Fanuc KAREL source: KC00004.KL

PROGRAM KC00004
%NOLOCKGROUP
%ENVIRONMENT PC
VAR
  I: INTEGER
  J: INTEGER
  K: INTEGER
  R: REAL
  B: BOOLEAN
  S: STRING[80]
  T: STRING[80]
  P: PATH
  Q: PATH
  AI: ARRAY[8] OF INTEGER
  AB: ARRAY[244] OF BYTE
BEGIN
  ADD_STRINGPC(AB,I,S,K)
END KC00004
